// TIA Portal V21 export
FUNCTION_BLOCK "ClassicLad"   // FB10, LAD
TITLE = ClassicLad
// Ladder on a classic CPU, with global tags.
   VAR_INPUT
      enable : Bool;
   END_VAR
   VAR_OUTPUT
      running : Bool;
   END_VAR
   VAR
      latched : Bool;
   END_VAR
BEGIN

REGION Network 1: Run the motor
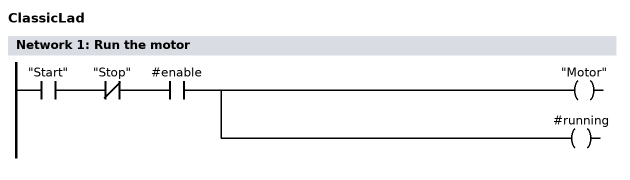
   RUNG wire#powerrail
      Contact( "Start" )
      I_Contact( "Stop" )
      Contact( #enable )
      wire#w1
      Coil( "Motor" )
   END_RUNG
   RUNG wire#w1
      Coil( #running )
   END_RUNG
   // the same network as SCL:
   "Motor" := "Start" AND NOT "Stop" AND #enable;
   #running := "Motor";
END_REGION
END_FUNCTION_BLOCK
